(*
    Organizes parsing and composing of XML data. Data can be treated as STRING or char array.
    Buffer size of file can be set via GVL_Param_TcUnit (xUnitBufferSize)
*)
FUNCTION_BLOCK FB_XmlControl
VAR
    XmlBuffer : FB_StreamBuffer;
    TagListBuffer : FB_StreamBuffer;
    Tags : T_MaxString;
    TagListSeekBuffer : FB_StreamBuffer;
    TagsSeek : STRING;
    TagBuffer : FB_StreamBuffer;
    Tag : T_MaxString;
    TagOpen: BOOL;
    Select : UDINT;
    SearchPosition : UDINT; 
END_VAR
VAR CONSTANT
    TAG_OPEN : STRING(1) := '<';
    TAG_CLOSE : STRING(1) := '>';
    END_TAG_CLOSE : STRING(2) := '/>';
    SPACE : STRING(1) := ' ';
    EQUALS : STRING(1) := '=';
    QUOTE : STRING(1) := '"';
    BACK_SLASH : STRING(1) := '\';
    FORWARD_SLASH : STRING(1) := '/';
    OPEN_COMMENT : STRING(5) := '<!-- ';
    CLOSE_COMMENT : STRING(4) := ' -->';
    TAB : STRING(2) := '$T';
    CR_LF : STRING(4) := '$R$N';

    // $OD : ASCII code for carriage return (CR)
    // $$ : to add a $R
    // $' : to add ' (apostrophe)
    // $L or $l : line feed
    // $N or $n : new line
    // $P or $p : next page
    // $R or $r : end of line
END_VAR

// Clears the contents of the entire buffer.
METHOD PUBLIC ClearBuffer
SearchPosition := 0;
TagListSeekBuffer.Length := 0;
XmlBuffer.Length := 0;
TagsSeek := '';
Tag := '';
END_METHOD

(*
    Closes a Tag:
    XML: <MyTag />'

    Method: XML.CloseTag();
*)
METHOD PUBLIC CloseTag : T_MaxString
VAR
    ClosedTag : T_MaxString;
END_VAR
IF TagOpen THEN
    XmlBuffer.Append := END_TAG_CLOSE;
    Select := TagListBuffer.FindBack(SearchString := FORWARD_SLASH);
    ClosedTag := TagListBuffer.CutOff(StartPos := Select);
    TagOpen := FALSE;
ELSE
    Select := TagListBuffer.FindBack(SearchString := FORWARD_SLASH);
    ClosedTag := TagListBuffer.CutOff(StartPos := Select);
    XmlBuffer.Append := TAG_OPEN;
    XmlBuffer.Append := ClosedTag;
    XmlBuffer.Append := TAG_CLOSE;
END_IF

CloseTag := ClosedTag;
END_METHOD

PROPERTY Length : UDINT
GET
Length := XmlBuffer.Length;
END_GET
END_PROPERTY

(*
    Adds a comment
    XML: <!-- MyComment -->

    XML.NewComment(Comment: = 'MyComment');
*)
METHOD PUBLIC NewComment
VAR_INPUT
    Comment : T_MaxString;
END_VAR
IF TagOpen THEN
    XmlBuffer.Append := TAG_CLOSE;
    TagOpen := FALSE;
END_IF;
XmlBuffer.Append := OPEN_COMMENT;
XmlBuffer.Append := Comment;
XmlBuffer.Append := CLOSE_COMMENT;
END_METHOD

(*
    Must be called after opening a new tag

    XML.NewParameter(Name: = 'ParaName', Value: = 'Value');
*)
METHOD PUBLIC NewParameter
VAR_INPUT
    Name : T_MaxString;
    Value : T_MaxString;
END_VAR
VAR
    ValueBytes : POINTER TO BYTE;
    ChunkBytes : POINTER TO BYTE;
    Chunk : T_MaxString;
    ChunkLength : INT;
    ValueLength : INT;
    Index : INT;
    Entity : STRING(6);
END_VAR
VAR CONSTANT
    AMPERSAND_BYTE : BYTE := 16#26;
    LESS_THAN_BYTE : BYTE := 16#3C;
    GREATER_THAN_BYTE : BYTE := 16#3E;
    QUOTE_BYTE : BYTE := 16#22;
    MAX_CHUNK_LENGTH : INT := 255;
END_VAR
XmlBuffer.Append := SPACE;
XmlBuffer.Append := Name;
XmlBuffer.Append := EQUALS;
XmlBuffer.Append := QUOTE;
(* The value is escaped: failure messages and skip reasons may contain characters that would end the
   attribute or start markup. Unescaped runs are appended in chunks, each entity on its own. *)
ValueBytes := ADR(Value);
ChunkBytes := ADR(Chunk);
ChunkLength := 0;
ValueLength := LEN(Value);
FOR Index := 0 TO ValueLength - 1 DO
    IF ValueBytes[Index] = AMPERSAND_BYTE THEN
        Entity := '&amp;';
    ELSIF ValueBytes[Index] = LESS_THAN_BYTE THEN
        Entity := '&lt;';
    ELSIF ValueBytes[Index] = GREATER_THAN_BYTE THEN
        Entity := '&gt;';
    ELSIF ValueBytes[Index] = QUOTE_BYTE THEN
        Entity := '&quot;';
    ELSE
        Entity := '';
        ChunkBytes[ChunkLength] := ValueBytes[Index];
        ChunkLength := ChunkLength + 1;
    END_IF
    IF LEN(Entity) > 0 OR ChunkLength >= MAX_CHUNK_LENGTH THEN
        ChunkBytes[ChunkLength] := 0;
        XmlBuffer.Append := Chunk;
        ChunkLength := 0;
        IF LEN(Entity) > 0 THEN
            XmlBuffer.Append := Entity;
        END_IF
    END_IF
END_FOR
IF ChunkLength > 0 THEN
    ChunkBytes[ChunkLength] := 0;
    XmlBuffer.Append := Chunk;
END_IF
XmlBuffer.Append := QUOTE;
END_METHOD

(*
    Creates a new Tag:
    XML: <MyTag>

    XML.NewTag(Name: = 'MyTag');
*)
METHOD PUBLIC NewTag
VAR_INPUT
    Name : T_MaxString;
END_VAR
IF TagOpen THEN
    XmlBuffer.Append := TAG_CLOSE;
END_IF;
XmlBuffer.Append := TAG_OPEN;
XmlBuffer.Append := Name;
TagOpen := TRUE;
TagListBuffer.Append := FORWARD_SLASH;
TagListBuffer.Append := Name;
END_METHOD

METHOD PUBLIC NewTagData
VAR_INPUT
    Data : T_MaxString;
END_VAR
XmlBuffer.Append := TAG_CLOSE;
XmlBuffer.Append := Data;
TagOpen := FALSE;
END_METHOD

METHOD PUBLIC SetBuffer
VAR_INPUT
    PointerToBuffer : POINTER TO BYTE; // ADR(..)
    SizeOfBuffer : UDINT; // SIZEOF(..)
END_VAR
XmlBuffer.SetBuffer(PointerToBufferAddress:= PointerToBuffer, SizeOfBuffer := SizeOfBuffer);
TagListBuffer.SetBuffer(PointerToBufferAddress := ADR(Tags), SizeOfBuffer := SIZEOF(Tags));
TagListSeekBuffer.SetBuffer(PointerToBufferAddress := ADR(TagsSeek), SizeOfBuffer := SIZEOF(TagsSeek));
TagBuffer.SetBuffer(PointerToBufferAddress := ADR(Tag), SizeOfBuffer := SIZEOF(Tag));
END_METHOD

(*
    Jump to the beginning of the XML data
    XML.ToStartBuffer();
*)
METHOD PUBLIC ToStartBuffer
SearchPosition := 0;
TagListSeekBuffer.Length := 0;
TagsSeek := '';
Tag := '';
END_METHOD

(*
    Add your own preffered fileheader like:
    XML: <?xml version="1.0" encoding="UTF-8"?>
    
    Start with calling this method before appending any other tags!

    XML.WriteDocumentHeader('<?xml version="1.0" encoding="UTF-8"?>');
*)
METHOD PUBLIC WriteDocumentHeader
VAR_INPUT
    Header : T_MaxString;
END_VAR
XmlBuffer.Append := Header;
END_METHOD

END_FUNCTION_BLOCK

(* stored: Version 1.1.0.1
   POU FB_XmlControl: Id {f48b7de2-5c07-4763-a8be-3d8ab3c1f58c}, SpecialFunc None
   Method ClearBuffer: Id {651b4460-232e-47e8-95ba-ecea1541fbb9}
   Method CloseTag: Id {eedd2aac-2425-4325-8128-bfe1e984f3f7}
   Property Length: Id {4fdf30b6-5fe7-4452-ad0a-85e866e236d0}
   Get Get: Id {267105d4-b124-4c5c-a359-0434c4992afc}
   Method NewComment: Id {0f41fa45-b92e-4e7e-b2b3-ecb5d5918326}
   Method NewParameter: Id {60c10606-ff09-4f9b-a3dd-0b54d0f565c7}
   Method NewTag: Id {c44bdbda-725a-4943-a5cc-fa5ea9485541}
   Method NewTagData: Id {e4679d3f-10eb-47fd-936c-97e3aaaa3768}
   Method SetBuffer: Id {cbfaa6d5-eab9-48d0-a339-a8bf334e344e}
   Method ToStartBuffer: Id {cb065068-a6c8-48d5-8c1d-535a21365348}
   Method WriteDocumentHeader: Id {14bf2549-9e7d-451f-8ab5-fe662eb30712} *)
